Fanuc KAREL source: ka00227.KL

-- PROVISIONAL review KL for V940-1; original PC SHA256 b1c522be1ac6652d90ab46c5a8e5753471ba38d94f7ed681ad284aca98e605d7
-- Incomplete behavior may be omitted. Consult companion uncertainty JSON. Do not deploy.
PROGRAM KA00227
%NOLOCKGROUP
-- UNRESOLVED_DECL SRC type=001100
-- UNRESOLVED_DECL DST type=001100
BEGIN
  -- V9_ZERO_TABLE_METADATA_HINT layout=0002_ascii; no indexed target words; source/name/runtime held
  -- UNRESOLVED_PC offsets 5-20; opcodes 22,22,30
  -- UNRESOLVED_PC offsets 25-29; opcodes 7F
END KA00227
